Fanuc KAREL source: kb00103.KL

-- PROVISIONAL review KL for V770-1; original PC SHA256 38ddc0e37e345050fb355f8c1ecdbbc94ed34dc21e7779b5ffc36218399de032
-- Incomplete behavior may be omitted. Consult companion uncertainty JSON. Do not deploy.
PROGRAM KB00103
%NOLOCKGROUP
BEGIN
  -- UNRESOLVED_PC offsets 5-12; opcodes 9D,23
  -- UNRESOLVED_PC offsets 17-24; opcodes 9D,23
  -- UNRESOLVED_PC offsets 29-38; opcodes 3F,75
  -- UNRESOLVED_PC offsets 43-50; opcodes 9D,23
  -- UNRESOLVED_PC offsets 55-62; opcodes 9D,23
  -- UNRESOLVED_PC offsets 67-74; opcodes 9D,23
  -- UNRESOLVED_PC offsets 79-86; opcodes 9D,23
  -- UNRESOLVED_PC offsets 91-98; opcodes 9D,23
  -- UNRESOLVED_PC offsets 103-110; opcodes 9D,23
  -- UNRESOLVED_PC offsets 115-122; opcodes 9D,23
  -- UNRESOLVED_PC offsets 127-199; opcodes 27,22,22,22,2A,22,22,22,22,22,22,22,22,31
  -- UNRESOLVED_PC offsets 204-208; opcodes 7F
END KB00103
